// TIA Portal V15.1 export
FUNCTION_BLOCK "Burner"   // FB1, LAD
TITLE = Burner
{ S7_Optimized_Access := 'TRUE' }
VERSION : 0.1
// One burner, docs/التشغيل.md §2 and decisions/0006
// stored: AutoNumber false, IsIECCheckEnabled false, MemoryReserve 100, SetENOAutomatically False
   VAR_INPUT
      Auto : Bool;   // AUTO/MAN selector, 1 = AUTO
      StartPB : Bool;   // START push button (NO)
      StopOK : Bool;   // STOP push button (NC): 1 = released
      LevelOK : Bool;   // Tank LSL reached (C07a)
      RunFb : Bool;   // Burner RUN feedback
      Lockout : Bool;   // Burner lockout signal (C07e)
      Fuel : Bool;   // Fuel mode (BR02 Rfuel2, R-12); FALSE for BR01
      TeA : Int;   // Thermocouple A raw, 0.1 degC
      TeB : Int;   // Thermocouple B raw, 0.1 degC
      Use24h : Bool;   // 24 h forced stop enabled (C07h, BR01 only)
      EStopOK : Bool;   // Sys.EStopOK
      ResetPulse : Bool;   // Sys.ResetPulse
      FirstScan : Bool;   // Sys.FirstScan
      SP : Int;   // Par.SP_V
      HYST : Int;   // Par.HYST_V
      STG : Int;   // Par.STG_V
      TStart : Time;   // Par.TStart_V
   END_VAR
   VAR_OUTPUT
      HeatReq : Bool;   // Heat request TL / L (E1 / E3)
      Stage2 : Bool;   // 2nd stage TR / T2 (E2 / E4)
      State : Int;   // 0 IDLE, 1 STARTING, 2 RUNNING, 3 FAULT
      Enabled : Bool;   // START given and not taken back (B-01)
      Tmax : Int;   // Higher of the two thermocouples, 0.1 degC
      F_EStop : Bool;   // Fault C01
      F_TC : Bool;   // Fault C0xd thermocouple
      F_Lockout : Bool;   // Fault C0xe lockout
      F_NoStart : Bool;   // Fault C0xf failed to start
      F_RunLost : Bool;   // Fault C0xg stopped by itself
      F_RunWrong : Bool;   // Fault R-09 RUN without request
      ParPending : Bool;   // R-11 / D6 / 0007: a validated entry differs from its active copy
   END_VAR
   VAR
      StartEdge : Bool;
      StartMem : Bool;
      AutoChg : Bool;
      AutoMem : Bool;
      FuelChg : Bool;
      FuelMem : Bool;
      TcOkA : Bool;
      TcOkB : Bool;
      TcOk : Bool;
      TcBad : Bool;
      Demand : Bool;
      HeatNeed : Bool;
      Ready : Bool;
      Active : Bool;
      Pause24 : Bool;
      RunWrong : Bool;
      NoStart : Bool;
      PwrUpDone : Bool;
      TcSlow : Bool;
      SP_Act : Int;
      HYST_Act : Int;
      STG_Act : Int;
      TStart_Act : Time;
      TOn : Int;
      TStg : Int;
      TStgOff : Int;
      T_PwrUp : TON_TIME;
      T_TcBad : TON_TIME;
      T_24h : TON_TIME;
      T_Pause : TON_TIME;
      T_RunOff : TON_TIME;
      T_Start : TON_TIME;
   END_VAR
   VAR_TEMP   // added for the SCL form of the ladder/FBD networks
      _w1 : Bool;
   END_VAR
BEGIN

REGION Network 1: R-05 — START edge: not on first scan, only after seen released, STOP wins
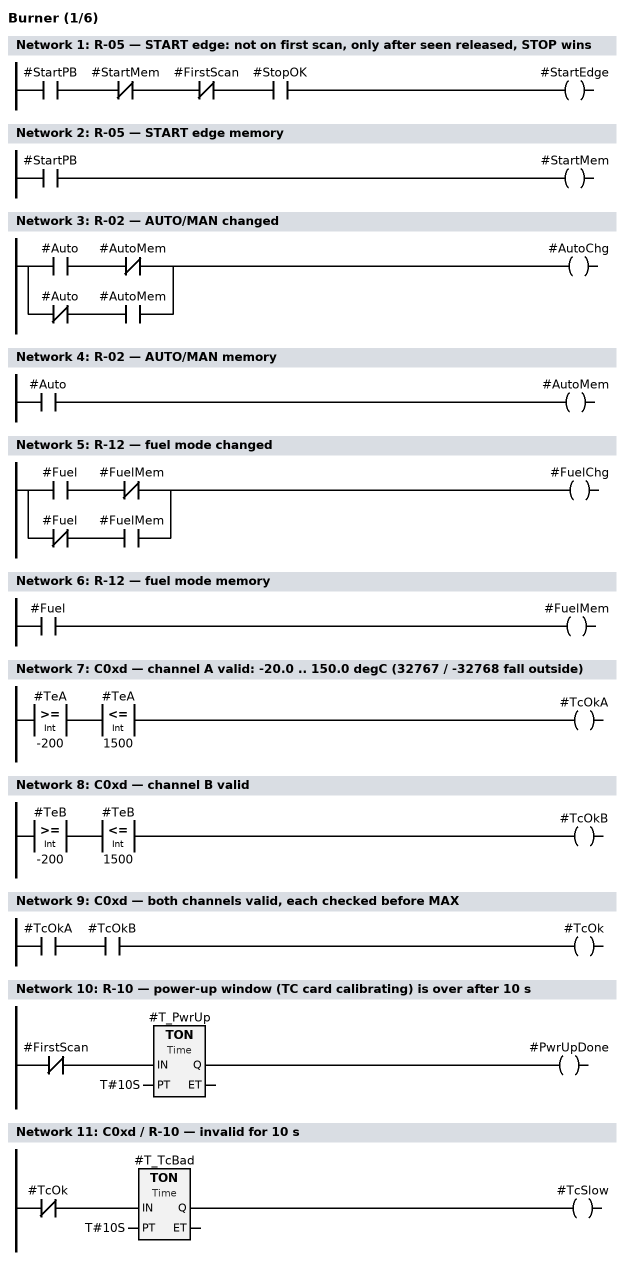
   RUNG wire#powerrail
      Contact( #StartPB )
      I_Contact( #StartMem )
      I_Contact( #FirstScan )
      Contact( #StopOK )
      Coil( #StartEdge )
   END_RUNG
   // the same network as SCL:
   #StartEdge := #StartPB AND NOT #StartMem AND NOT #FirstScan AND #StopOK;
END_REGION

REGION Network 2: R-05 — START edge memory
   RUNG wire#powerrail
      Contact( #StartPB )
      Coil( #StartMem )
   END_RUNG
   // the same network as SCL:
   #StartMem := #StartPB;
END_REGION

REGION Network 3: R-02 — AUTO/MAN changed
   RUNG wire#powerrail
      Contact( #Auto )
      I_Contact( #AutoMem )
      wire#w1
      Coil( #AutoChg )
   END_RUNG
   RUNG wire#powerrail
      I_Contact( #Auto )
      Contact( #AutoMem )
   END_RUNG wire#w1
   // the same network as SCL:
   #AutoChg := (#Auto AND NOT #AutoMem) OR (NOT #Auto AND #AutoMem);
END_REGION

REGION Network 4: R-02 — AUTO/MAN memory
   RUNG wire#powerrail
      Contact( #Auto )
      Coil( #AutoMem )
   END_RUNG
   // the same network as SCL:
   #AutoMem := #Auto;
END_REGION

REGION Network 5: R-12 — fuel mode changed
   RUNG wire#powerrail
      Contact( #Fuel )
      I_Contact( #FuelMem )
      wire#w1
      Coil( #FuelChg )
   END_RUNG
   RUNG wire#powerrail
      I_Contact( #Fuel )
      Contact( #FuelMem )
   END_RUNG wire#w1
   // the same network as SCL:
   #FuelChg := (#Fuel AND NOT #FuelMem) OR (NOT #Fuel AND #FuelMem);
END_REGION

REGION Network 6: R-12 — fuel mode memory
   RUNG wire#powerrail
      Contact( #Fuel )
      Coil( #FuelMem )
   END_RUNG
   // the same network as SCL:
   #FuelMem := #Fuel;
END_REGION

REGION Network 7: C0xd — channel A valid: -20.0 .. 150.0 degC (32767 / -32768 fall outside)
   RUNG wire#powerrail
      { S7_Templates := "SrcType := Int" } GE_Contact(in1 := #TeA, in2 := -200)
      { S7_Templates := "SrcType := Int" } LE_Contact(in1 := #TeA, in2 := 1500)
      Coil( #TcOkA )
   END_RUNG
   // the same network as SCL:
   #TcOkA := (#TeA >= (-200)) AND (#TeA <= 1500);
END_REGION

REGION Network 8: C0xd — channel B valid
   RUNG wire#powerrail
      { S7_Templates := "SrcType := Int" } GE_Contact(in1 := #TeB, in2 := -200)
      { S7_Templates := "SrcType := Int" } LE_Contact(in1 := #TeB, in2 := 1500)
      Coil( #TcOkB )
   END_RUNG
   // the same network as SCL:
   #TcOkB := (#TeB >= (-200)) AND (#TeB <= 1500);
END_REGION

REGION Network 9: C0xd — both channels valid, each checked before MAX
   RUNG wire#powerrail
      Contact( #TcOkA )
      Contact( #TcOkB )
      Coil( #TcOk )
   END_RUNG
   // the same network as SCL:
   #TcOk := #TcOkA AND #TcOkB;
END_REGION

REGION Network 10: R-10 — power-up window (TC card calibrating) is over after 10 s
   RUNG wire#powerrail
      I_Contact( #FirstScan )
      { S7_Templates := "time_type := Time" } #T_PwrUp.TON(pt := T#10S, et =>)
      Coil( #PwrUpDone )
   END_RUNG
   // the same network as SCL:
   #T_PwrUp(IN := NOT #FirstScan, PT := T#10S);   // TON
   #PwrUpDone := #T_PwrUp.Q;
END_REGION

REGION Network 11: C0xd / R-10 — invalid for 10 s
   RUNG wire#powerrail
      I_Contact( #TcOk )
      { S7_Templates := "time_type := Time" } #T_TcBad.TON(pt := T#10S, et =>)
      Coil( #TcSlow )
   END_RUNG
   // the same network as SCL:
   #T_TcBad(IN := NOT #TcOk, PT := T#10S);   // TON
   #TcSlow := #T_TcBad.Q;
END_REGION

REGION Network 12: C0xd / R-10 — invalid = fault: at once, or after 10 s right after power-up
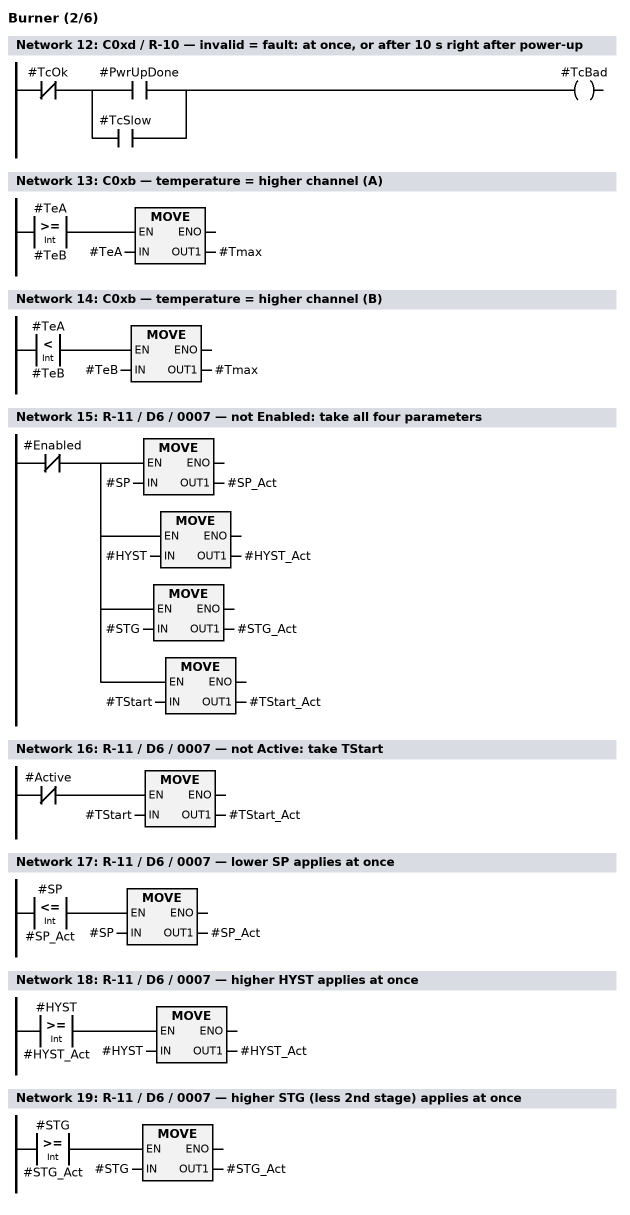
   RUNG wire#powerrail
      I_Contact( #TcOk )
      wire#w1
      Contact( #PwrUpDone )
      wire#w2
      Coil( #TcBad )
   END_RUNG
   RUNG wire#w1
      Contact( #TcSlow )
   END_RUNG wire#w2
   // the same network as SCL:
   #TcBad := NOT #TcOk AND (#PwrUpDone OR #TcSlow);
END_REGION

REGION Network 13: C0xb — temperature = higher channel (A)
   RUNG wire#powerrail
      { S7_Templates := "SrcType := Int" } GE_Contact(in1 := #TeA, in2 := #TeB)
      { S7_GenerateENO := "TRUE" } Move(in := #TeA, out1 => #Tmax)
   END_RUNG
   // the same network as SCL:
   IF #TeA >= #TeB THEN #Tmax := #TeA; END_IF;
END_REGION

REGION Network 14: C0xb — temperature = higher channel (B)
   RUNG wire#powerrail
      { S7_Templates := "SrcType := Int" } LT_Contact(in1 := #TeA, in2 := #TeB)
      { S7_GenerateENO := "TRUE" } Move(in := #TeB, out1 => #Tmax)
   END_RUNG
   // the same network as SCL:
   IF #TeA < #TeB THEN #Tmax := #TeB; END_IF;
END_REGION

REGION Network 15: R-11 / D6 / 0007 — not Enabled: take all four parameters
   RUNG wire#powerrail
      I_Contact( #Enabled )
      wire#w1
      { S7_GenerateENO := "TRUE" } Move(in := #SP, out1 => #SP_Act)
   END_RUNG
   RUNG wire#w1
      { S7_GenerateENO := "TRUE" } Move(in := #HYST, out1 => #HYST_Act)
   END_RUNG
   RUNG wire#w1
      { S7_GenerateENO := "TRUE" } Move(in := #STG, out1 => #STG_Act)
   END_RUNG
   RUNG wire#w1
      { S7_GenerateENO := "TRUE" } Move(in := #TStart, out1 => #TStart_Act)
   END_RUNG
   // the same network as SCL:
   IF NOT #Enabled THEN
       #SP_Act := #SP;
       #HYST_Act := #HYST;
       #STG_Act := #STG;
       #TStart_Act := #TStart;
   END_IF;
END_REGION

REGION Network 16: R-11 / D6 / 0007 — not Active: take TStart
   RUNG wire#powerrail
      I_Contact( #Active )
      { S7_GenerateENO := "TRUE" } Move(in := #TStart, out1 => #TStart_Act)
   END_RUNG
   // the same network as SCL:
   IF NOT #Active THEN #TStart_Act := #TStart; END_IF;
END_REGION

REGION Network 17: R-11 / D6 / 0007 — lower SP applies at once
   RUNG wire#powerrail
      { S7_Templates := "SrcType := Int" } LE_Contact(in1 := #SP, in2 := #SP_Act)
      { S7_GenerateENO := "TRUE" } Move(in := #SP, out1 => #SP_Act)
   END_RUNG
   // the same network as SCL:
   IF #SP <= #SP_Act THEN #SP_Act := #SP; END_IF;
END_REGION

REGION Network 18: R-11 / D6 / 0007 — higher HYST applies at once
   RUNG wire#powerrail
      { S7_Templates := "SrcType := Int" } GE_Contact(in1 := #HYST, in2 := #HYST_Act)
      { S7_GenerateENO := "TRUE" } Move(in := #HYST, out1 => #HYST_Act)
   END_RUNG
   // the same network as SCL:
   IF #HYST >= #HYST_Act THEN #HYST_Act := #HYST; END_IF;
END_REGION

REGION Network 19: R-11 / D6 / 0007 — higher STG (less 2nd stage) applies at once
   RUNG wire#powerrail
      { S7_Templates := "SrcType := Int" } GE_Contact(in1 := #STG, in2 := #STG_Act)
      { S7_GenerateENO := "TRUE" } Move(in := #STG, out1 => #STG_Act)
   END_RUNG
   // the same network as SCL:
   IF #STG >= #STG_Act THEN #STG_Act := #STG; END_IF;
END_REGION

REGION Network 20: R-11 / D6 / 0007 — pending while any entry differs from its active copy
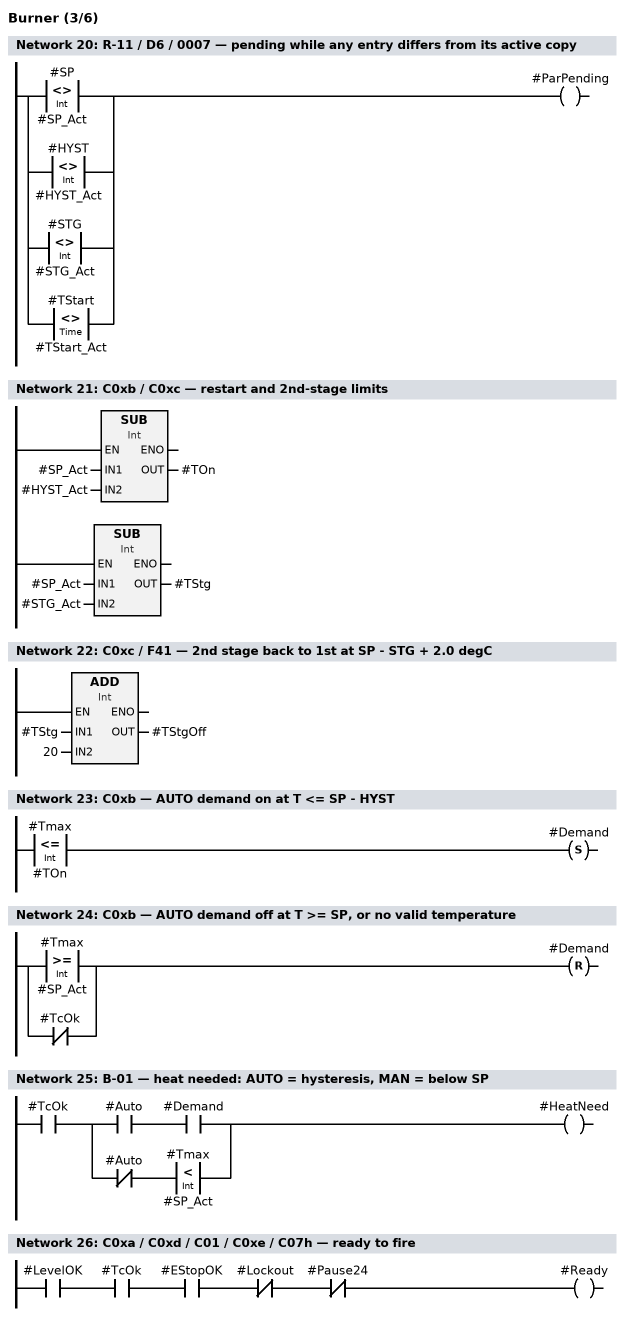
   RUNG wire#powerrail
      { S7_Templates := "SrcType := Int" } NE_Contact(in1 := #SP, in2 := #SP_Act)
      wire#w1
      Coil( #ParPending )
   END_RUNG
   RUNG wire#powerrail
      { S7_Templates := "SrcType := Int" } NE_Contact(in1 := #HYST, in2 := #HYST_Act)
   END_RUNG wire#w1
   RUNG wire#powerrail
      { S7_Templates := "SrcType := Int" } NE_Contact(in1 := #STG, in2 := #STG_Act)
   END_RUNG wire#w1
   RUNG wire#powerrail
      { S7_Templates := "SrcType := Time" } NE_Contact(in1 := #TStart, in2 := #TStart_Act)
   END_RUNG wire#w1
   // the same network as SCL:
   #ParPending := (#SP <> #SP_Act) OR (#HYST <> #HYST_Act) OR (#STG <> #STG_Act) OR (#TStart <> #TStart_Act);
END_REGION

REGION Network 21: C0xb / C0xc — restart and 2nd-stage limits
   RUNG wire#powerrail
      { S7_Templates := "SrcType := Int"; S7_GenerateENO := "TRUE" } Sub(in1 := #SP_Act, in2 := #HYST_Act, out => #TOn)
   END_RUNG
   RUNG wire#powerrail
      { S7_Templates := "SrcType := Int"; S7_GenerateENO := "TRUE" } Sub(in1 := #SP_Act, in2 := #STG_Act, out => #TStg)
   END_RUNG
   // the same network as SCL:
   #TOn := #SP_Act - #HYST_Act;
   #TStg := #SP_Act - #STG_Act;
END_REGION

REGION Network 22: C0xc / F41 — 2nd stage back to 1st at SP - STG + 2.0 degC
   RUNG wire#powerrail
      { S7_Templates := "SrcType := Int"; S7_GenerateENO := "TRUE" } Add(in1 := #TStg, in2 := 20, out => #TStgOff)
   END_RUNG
   // the same network as SCL:
   #TStgOff := #TStg + 20;
END_REGION

REGION Network 23: C0xb — AUTO demand on at T <= SP - HYST
   RUNG wire#powerrail
      { S7_Templates := "SrcType := Int" } LE_Contact(in1 := #Tmax, in2 := #TOn)
      S_Coil( #Demand )
   END_RUNG
   // the same network as SCL:
   IF #Tmax <= #TOn THEN #Demand := TRUE; END_IF;
END_REGION

REGION Network 24: C0xb — AUTO demand off at T >= SP, or no valid temperature
   RUNG wire#powerrail
      { S7_Templates := "SrcType := Int" } GE_Contact(in1 := #Tmax, in2 := #SP_Act)
      wire#w1
      R_Coil( #Demand )
   END_RUNG
   RUNG wire#powerrail
      I_Contact( #TcOk )
   END_RUNG wire#w1
   // the same network as SCL:
   IF (#Tmax >= #SP_Act) OR NOT #TcOk THEN #Demand := FALSE; END_IF;
END_REGION

REGION Network 25: B-01 — heat needed: AUTO = hysteresis, MAN = below SP
   RUNG wire#powerrail
      Contact( #TcOk )
      wire#w1
      Contact( #Auto )
      Contact( #Demand )
      wire#w2
      Coil( #HeatNeed )
   END_RUNG
   RUNG wire#w1
      I_Contact( #Auto )
      { S7_Templates := "SrcType := Int" } LT_Contact(in1 := #Tmax, in2 := #SP_Act)
   END_RUNG wire#w2
   // the same network as SCL:
   #HeatNeed := #TcOk AND ((#Auto AND #Demand) OR (NOT #Auto AND (#Tmax < #SP_Act)));
END_REGION

REGION Network 26: C0xa / C0xd / C01 / C0xe / C07h — ready to fire
   RUNG wire#powerrail
      Contact( #LevelOK )
      Contact( #TcOk )
      Contact( #EStopOK )
      I_Contact( #Lockout )
      I_Contact( #Pause24 )
      Coil( #Ready )
   END_RUNG
   // the same network as SCL:
   #Ready := #LevelOK AND #TcOk AND #EStopOK AND NOT #Lockout AND NOT #Pause24;
END_REGION

REGION Network 27: C07h / R-08 — 24 h of continuous request: forced stop
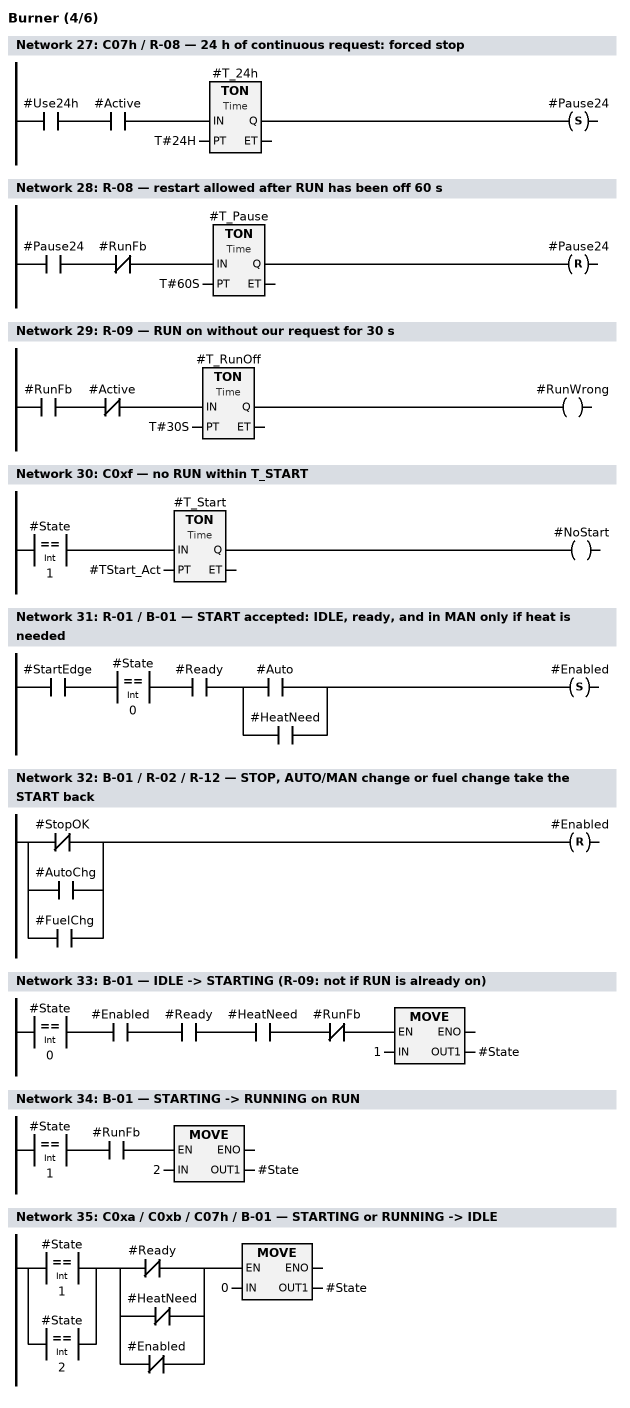
   RUNG wire#powerrail
      Contact( #Use24h )
      Contact( #Active )
      { S7_Templates := "time_type := Time" } #T_24h.TON(pt := T#24H, et =>)
      S_Coil( #Pause24 )
   END_RUNG
   // the same network as SCL:
   #T_24h(IN := #Use24h AND #Active, PT := T#24H);   // TON
   IF #T_24h.Q THEN #Pause24 := TRUE; END_IF;
END_REGION

REGION Network 28: R-08 — restart allowed after RUN has been off 60 s
   RUNG wire#powerrail
      Contact( #Pause24 )
      I_Contact( #RunFb )
      { S7_Templates := "time_type := Time" } #T_Pause.TON(pt := T#60S, et =>)
      R_Coil( #Pause24 )
   END_RUNG
   // the same network as SCL:
   #T_Pause(IN := #Pause24 AND NOT #RunFb, PT := T#60S);   // TON
   IF #T_Pause.Q THEN #Pause24 := FALSE; END_IF;
END_REGION

REGION Network 29: R-09 — RUN on without our request for 30 s
   RUNG wire#powerrail
      Contact( #RunFb )
      I_Contact( #Active )
      { S7_Templates := "time_type := Time" } #T_RunOff.TON(pt := T#30S, et =>)
      Coil( #RunWrong )
   END_RUNG
   // the same network as SCL:
   #T_RunOff(IN := #RunFb AND NOT #Active, PT := T#30S);   // TON
   #RunWrong := #T_RunOff.Q;
END_REGION

REGION Network 30: C0xf — no RUN within T_START
   RUNG wire#powerrail
      { S7_Templates := "SrcType := Int" } EQ_Contact(in1 := #State, in2 := 1)
      { S7_Templates := "time_type := Time" } #T_Start.TON(pt := #TStart_Act, et =>)
      Coil( #NoStart )
   END_RUNG
   // the same network as SCL:
   #T_Start(IN := #State = 1, PT := #TStart_Act);   // TON
   #NoStart := #T_Start.Q;
END_REGION

REGION Network 31: R-01 / B-01 — START accepted: IDLE, ready, and in MAN only if heat is needed
   RUNG wire#powerrail
      Contact( #StartEdge )
      { S7_Templates := "SrcType := Int" } EQ_Contact(in1 := #State, in2 := 0)
      Contact( #Ready )
      wire#w1
      Contact( #Auto )
      wire#w2
      S_Coil( #Enabled )
   END_RUNG
   RUNG wire#w1
      Contact( #HeatNeed )
   END_RUNG wire#w2
   // the same network as SCL:
   IF #StartEdge AND (#State = 0) AND #Ready AND (#Auto OR #HeatNeed) THEN #Enabled := TRUE; END_IF;
END_REGION

REGION Network 32: B-01 / R-02 / R-12 — STOP, AUTO/MAN change or fuel change take the START back
   RUNG wire#powerrail
      I_Contact( #StopOK )
      wire#w1
      R_Coil( #Enabled )
   END_RUNG
   RUNG wire#powerrail
      Contact( #AutoChg )
   END_RUNG wire#w1
   RUNG wire#powerrail
      Contact( #FuelChg )
   END_RUNG wire#w1
   // the same network as SCL:
   IF NOT #StopOK OR #AutoChg OR #FuelChg THEN #Enabled := FALSE; END_IF;
END_REGION

REGION Network 33: B-01 — IDLE -> STARTING (R-09: not if RUN is already on)
   RUNG wire#powerrail
      { S7_Templates := "SrcType := Int" } EQ_Contact(in1 := #State, in2 := 0)
      Contact( #Enabled )
      Contact( #Ready )
      Contact( #HeatNeed )
      I_Contact( #RunFb )
      { S7_GenerateENO := "TRUE" } Move(in := 1, out1 => #State)
   END_RUNG
   // the same network as SCL:
   IF (#State = 0) AND #Enabled AND #Ready AND #HeatNeed AND NOT #RunFb THEN #State := 1; END_IF;
END_REGION

REGION Network 34: B-01 — STARTING -> RUNNING on RUN
   RUNG wire#powerrail
      { S7_Templates := "SrcType := Int" } EQ_Contact(in1 := #State, in2 := 1)
      Contact( #RunFb )
      { S7_GenerateENO := "TRUE" } Move(in := 2, out1 => #State)
   END_RUNG
   // the same network as SCL:
   IF (#State = 1) AND #RunFb THEN #State := 2; END_IF;
END_REGION

REGION Network 35: C0xa / C0xb / C07h / B-01 — STARTING or RUNNING -> IDLE
   RUNG wire#powerrail
      { S7_Templates := "SrcType := Int" } EQ_Contact(in1 := #State, in2 := 1)
      wire#w1
      I_Contact( #Ready )
      wire#w2
      { S7_GenerateENO := "TRUE" } Move(in := 0, out1 => #State)
   END_RUNG
   RUNG wire#powerrail
      { S7_Templates := "SrcType := Int" } EQ_Contact(in1 := #State, in2 := 2)
   END_RUNG wire#w1
   RUNG wire#w1
      I_Contact( #HeatNeed )
   END_RUNG wire#w2
   RUNG wire#w1
      I_Contact( #Enabled )
   END_RUNG wire#w2
   // the same network as SCL:
   IF ((#State = 1) OR (#State = 2)) AND (NOT #Ready OR NOT #HeatNeed OR NOT #Enabled) THEN
       #State := 0;
   END_IF;
END_REGION

REGION Network 36: R-03 — MAN: one cycle; any stop needs a new START
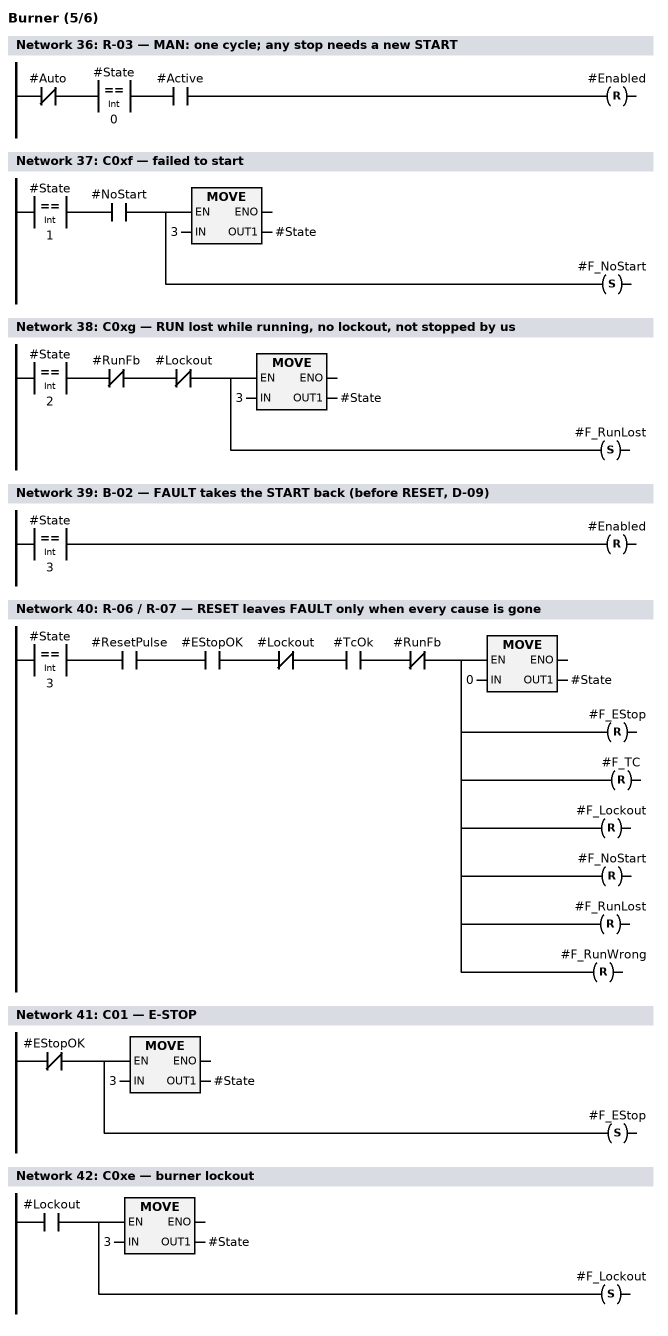
   RUNG wire#powerrail
      I_Contact( #Auto )
      { S7_Templates := "SrcType := Int" } EQ_Contact(in1 := #State, in2 := 0)
      Contact( #Active )
      R_Coil( #Enabled )
   END_RUNG
   // the same network as SCL:
   IF NOT #Auto AND (#State = 0) AND #Active THEN #Enabled := FALSE; END_IF;
END_REGION

REGION Network 37: C0xf — failed to start
   RUNG wire#powerrail
      { S7_Templates := "SrcType := Int" } EQ_Contact(in1 := #State, in2 := 1)
      Contact( #NoStart )
      wire#w1
      { S7_GenerateENO := "TRUE" } Move(in := 3, out1 => #State)
   END_RUNG
   RUNG wire#w1
      S_Coil( #F_NoStart )
   END_RUNG
   // the same network as SCL:
   #_w1 := (#State = 1) AND #NoStart;
   IF #_w1 THEN
       #State := 3;
       #F_NoStart := TRUE;
   END_IF;
END_REGION

REGION Network 38: C0xg — RUN lost while running, no lockout, not stopped by us
   RUNG wire#powerrail
      { S7_Templates := "SrcType := Int" } EQ_Contact(in1 := #State, in2 := 2)
      I_Contact( #RunFb )
      I_Contact( #Lockout )
      wire#w1
      { S7_GenerateENO := "TRUE" } Move(in := 3, out1 => #State)
   END_RUNG
   RUNG wire#w1
      S_Coil( #F_RunLost )
   END_RUNG
   // the same network as SCL:
   #_w1 := (#State = 2) AND NOT #RunFb AND NOT #Lockout;
   IF #_w1 THEN
       #State := 3;
       #F_RunLost := TRUE;
   END_IF;
END_REGION

REGION Network 39: B-02 — FAULT takes the START back (before RESET, D-09)
   RUNG wire#powerrail
      { S7_Templates := "SrcType := Int" } EQ_Contact(in1 := #State, in2 := 3)
      R_Coil( #Enabled )
   END_RUNG
   // the same network as SCL:
   IF #State = 3 THEN #Enabled := FALSE; END_IF;
END_REGION

REGION Network 40: R-06 / R-07 — RESET leaves FAULT only when every cause is gone
   RUNG wire#powerrail
      { S7_Templates := "SrcType := Int" } EQ_Contact(in1 := #State, in2 := 3)
      Contact( #ResetPulse )
      Contact( #EStopOK )
      I_Contact( #Lockout )
      Contact( #TcOk )
      I_Contact( #RunFb )
      wire#w1
      { S7_GenerateENO := "TRUE" } Move(in := 0, out1 => #State)
   END_RUNG
   RUNG wire#w1
      R_Coil( #F_EStop )
   END_RUNG
   RUNG wire#w1
      R_Coil( #F_TC )
   END_RUNG
   RUNG wire#w1
      R_Coil( #F_Lockout )
   END_RUNG
   RUNG wire#w1
      R_Coil( #F_NoStart )
   END_RUNG
   RUNG wire#w1
      R_Coil( #F_RunLost )
   END_RUNG
   RUNG wire#w1
      R_Coil( #F_RunWrong )
   END_RUNG
   // the same network as SCL:
   #_w1 := (#State = 3) AND #ResetPulse AND #EStopOK AND NOT #Lockout AND #TcOk AND NOT #RunFb;
   IF #_w1 THEN
       #State := 0;
       #F_EStop := FALSE;
       #F_TC := FALSE;
       #F_Lockout := FALSE;
       #F_NoStart := FALSE;
       #F_RunLost := FALSE;
       #F_RunWrong := FALSE;
   END_IF;
END_REGION

REGION Network 41: C01 — E-STOP
   RUNG wire#powerrail
      I_Contact( #EStopOK )
      wire#w1
      { S7_GenerateENO := "TRUE" } Move(in := 3, out1 => #State)
   END_RUNG
   RUNG wire#w1
      S_Coil( #F_EStop )
   END_RUNG
   // the same network as SCL:
   IF NOT #EStopOK THEN
       #State := 3;
       #F_EStop := TRUE;
   END_IF;
END_REGION

REGION Network 42: C0xe — burner lockout
   RUNG wire#powerrail
      Contact( #Lockout )
      wire#w1
      { S7_GenerateENO := "TRUE" } Move(in := 3, out1 => #State)
   END_RUNG
   RUNG wire#w1
      S_Coil( #F_Lockout )
   END_RUNG
   // the same network as SCL:
   IF #Lockout THEN
       #State := 3;
       #F_Lockout := TRUE;
   END_IF;
END_REGION

REGION Network 43: C0xd — thermocouple fault
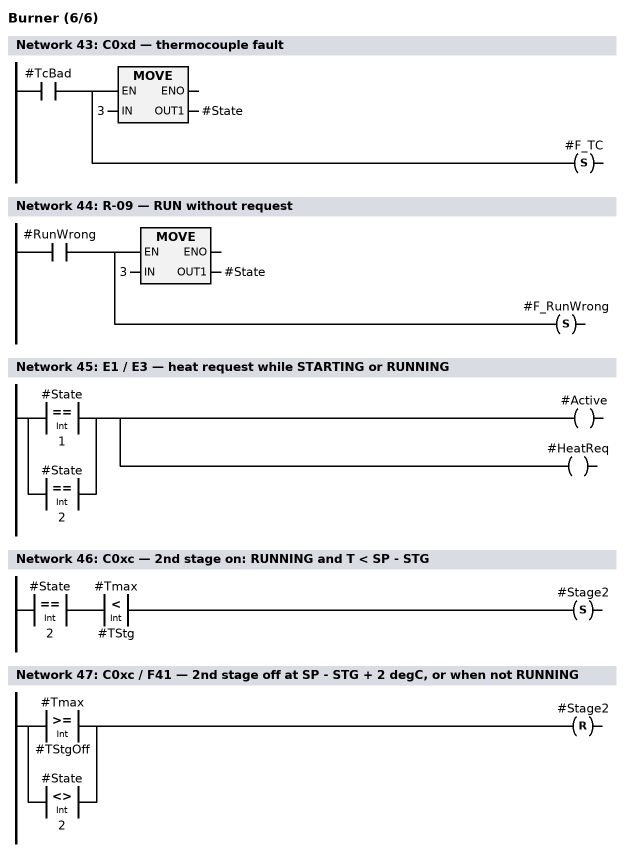
   RUNG wire#powerrail
      Contact( #TcBad )
      wire#w1
      { S7_GenerateENO := "TRUE" } Move(in := 3, out1 => #State)
   END_RUNG
   RUNG wire#w1
      S_Coil( #F_TC )
   END_RUNG
   // the same network as SCL:
   IF #TcBad THEN
       #State := 3;
       #F_TC := TRUE;
   END_IF;
END_REGION

REGION Network 44: R-09 — RUN without request
   RUNG wire#powerrail
      Contact( #RunWrong )
      wire#w1
      { S7_GenerateENO := "TRUE" } Move(in := 3, out1 => #State)
   END_RUNG
   RUNG wire#w1
      S_Coil( #F_RunWrong )
   END_RUNG
   // the same network as SCL:
   IF #RunWrong THEN
       #State := 3;
       #F_RunWrong := TRUE;
   END_IF;
END_REGION

REGION Network 45: E1 / E3 — heat request while STARTING or RUNNING
   RUNG wire#powerrail
      { S7_Templates := "SrcType := Int" } EQ_Contact(in1 := #State, in2 := 1)
      wire#w1
      Coil( #Active )
   END_RUNG
   RUNG wire#powerrail
      { S7_Templates := "SrcType := Int" } EQ_Contact(in1 := #State, in2 := 2)
   END_RUNG wire#w1
   RUNG wire#w1
      Coil( #HeatReq )
   END_RUNG
   // the same network as SCL:
   #Active := (#State = 1) OR (#State = 2);
   #HeatReq := #Active;
END_REGION

REGION Network 46: C0xc — 2nd stage on: RUNNING and T < SP - STG
   RUNG wire#powerrail
      { S7_Templates := "SrcType := Int" } EQ_Contact(in1 := #State, in2 := 2)
      { S7_Templates := "SrcType := Int" } LT_Contact(in1 := #Tmax, in2 := #TStg)
      S_Coil( #Stage2 )
   END_RUNG
   // the same network as SCL:
   IF (#State = 2) AND (#Tmax < #TStg) THEN #Stage2 := TRUE; END_IF;
END_REGION

REGION Network 47: C0xc / F41 — 2nd stage off at SP - STG + 2 degC, or when not RUNNING
   RUNG wire#powerrail
      { S7_Templates := "SrcType := Int" } GE_Contact(in1 := #Tmax, in2 := #TStgOff)
      wire#w1
      R_Coil( #Stage2 )
   END_RUNG
   RUNG wire#powerrail
      { S7_Templates := "SrcType := Int" } NE_Contact(in1 := #State, in2 := 2)
   END_RUNG wire#w1
   // the same network as SCL:
   IF (#Tmax >= #TStgOff) OR (#State <> 2) THEN #Stage2 := FALSE; END_IF;
END_REGION
END_FUNCTION_BLOCK
